FUNCTION_BLOCK Controle_Revezamento_2 (* Revezamento de 2 equipamentos por tempo como principal (mesmo padrao do Controle_Revezamento_3) *)
  (* Standard: 61499-2 *)
  (* Version 1.0, 21/10/2026, Hidryco, Hidryco, 1.0: Revezamento de 2 equipamentos por tempo como principal (mesmo padrao do Controle_Revezamento_3) *)
  PACKAGE Hidryco.HidrycoLib;
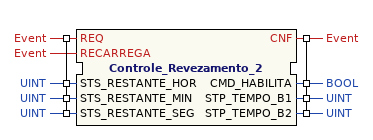
  EVENT_INPUT
    REQ WITH STS_RESTANTE_HOR, STS_RESTANTE_MIN, STS_RESTANTE_SEG; (* Status vindo do processo *)
    RECARREGA; (* Reenvia os ajustes persistentes (chamado no fim do INIT do processo) *)
  END_EVENT
  EVENT_OUTPUT
    CNF WITH CMD_HABILITA, STP_TEMPO_B1, STP_TEMPO_B2; (* Ajustes para o processo (mudanca na IHM, OPC UA ou recarga) *)
  END_EVENT
  VAR_INPUT
    STS_RESTANTE_HOR : UINT; (* Tempo para a troca da principal (h) *)
    STS_RESTANTE_MIN : UINT; (* Tempo para a troca da principal (min) *)
    STS_RESTANTE_SEG : UINT; (* Tempo para a troca da principal (s) *)
  END_VAR
  VAR_OUTPUT
    CMD_HABILITA : BOOL; (* Troca da principal por tempo *)
    STP_TEMPO_B1 : UINT; (* Horas do equipamento 1 como principal *)
    STP_TEMPO_B2 : UINT; (* Horas do equipamento 2 como principal *)
  END_VAR
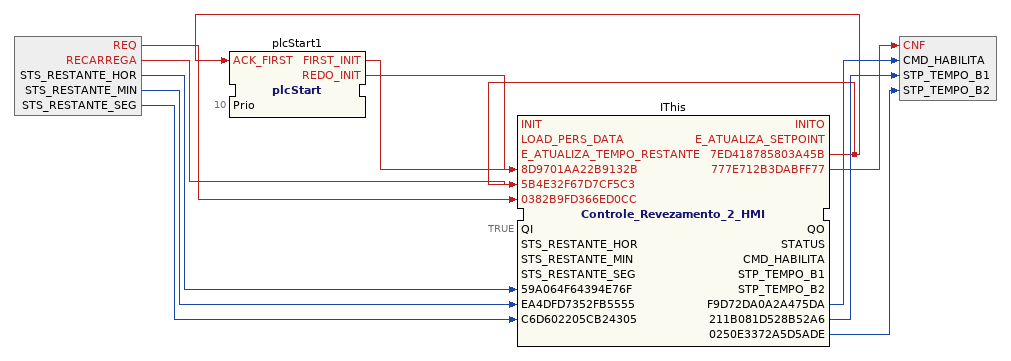
  FBS
    IThis : Controle_Revezamento_2_HMI(QI := TRUE);
    plcStart1 : plcStart(Prio := 10);
  END_FBS
  EVENT_CONNECTIONS
    plcStart1.FIRST_INIT TO IThis.8D9701AA22B9132B;
    plcStart1.REDO_INIT TO IThis.8D9701AA22B9132B;
    IThis.7ED418785803A45B TO IThis.5B4E32F67D7CF5C3;
    IThis.7ED418785803A45B TO plcStart1.ACK_FIRST;
    RECARREGA TO IThis.5B4E32F67D7CF5C3;
    IThis.777E712B3DABFF77 TO CNF;
    REQ TO IThis.0382B9FD366ED0CC;
  END_CONNECTIONS
  DATA_CONNECTIONS
    IThis.F9D72DA0A2A475DA TO CMD_HABILITA;
    IThis.211B081D528B52A6 TO STP_TEMPO_B1;
    IThis.0250E3372A5D5ADE TO STP_TEMPO_B2;
    STS_RESTANTE_HOR TO IThis.59A064F64394E76F;
    STS_RESTANTE_MIN TO IThis.EA4DFD7352FB5555;
    STS_RESTANTE_SEG TO IThis.C6D602205CB24305;
  END_CONNECTIONS
END_FUNCTION_BLOCK
